Fanuc TP program (LS listing): THREADPROG.LS

/PROG  THREADPROG
/ATTR
OWNER		= MNEDITOR;
COMMENT		= "RoboDK sequence";
PROG_SIZE	= 0;
CREATE		= DATE 26-10-26  TIME 01:01:16;
MODIFIED	= DATE 26-10-26  TIME 01:01:16;
FILE_NAME	= ;
VERSION	= 0;
LINE_COUNT	= 2;
MEMORY_SIZE	= 0;
PROTECT		= READ_WRITE;
TCD:  STACK_SIZE	= 0,
      TASK_PRIORITY	= 50,
TIME_SLICE	= 0,
BUSY_LAMP_OFF	= 0,
ABORT_REQUEST	= 0,
PAUSE_REQUEST	= 0;
DEFAULT_GROUP	= 1,*,*,*,*;
CONTROL_CODE	= 00000000 00000000;
/MN
   1:  UTOOL_NUM=1;
   2:  UFRAME_NUM=1;
/POS
/END
